(* IEC 61131-3 sources: trust-platform/examples/OSCAT/greenhouse_temperature/non-oop/src, 3 files *)

(* ---- Configuration.st ---- *)
CONFIGURATION GreenhouseTemperatureClassicConfiguration
RESOURCE Cpu0 ON PLC
    TASK MainTask (INTERVAL := T#100ms, PRIORITY := 1);
    PROGRAM Main WITH MainTask : Main;
END_RESOURCE
END_CONFIGURATION

(* ---- Main.st ---- *)
PROGRAM Main
VAR
    TemperatureConversion : TEMPERATURE;
    VentilationSwitch : HYST;
    TemperatureCelsius : REAL := REAL#29.0;
    TemperatureKelvin : REAL;
    TemperatureFahrenheit : REAL;
    VentilationRequest : BOOL;
END_VAR

TemperatureConversion(C := TemperatureCelsius);
TemperatureKelvin := TemperatureConversion.YK;
TemperatureFahrenheit := TemperatureConversion.YF;
VentilationSwitch(In := TemperatureCelsius, HIGH_LIMIT := REAL#28.0, LOW_LIMIT := REAL#18.0);
VentilationRequest := VentilationSwitch.Q;
END_PROGRAM

(* ---- Tests.st ---- *)
TEST_PROGRAM GreenhouseTemperatureClassicConvertsAndRequestsVentilation
VAR
    TemperatureConversion : TEMPERATURE;
    VentilationSwitch : HYST;
END_VAR

TemperatureConversion(C := REAL#29.0);
VentilationSwitch(In := REAL#29.0, HIGH_LIMIT := REAL#28.0, LOW_LIMIT := REAL#18.0);

ASSERT_NEAR(EXPECTED := REAL#302.15, ACTUAL := TemperatureConversion.YK, DELTA := REAL#0.01);
ASSERT_TRUE(IN := VentilationSwitch.Q);
END_TEST_PROGRAM
